FUNCTION_BLOCK "FB_ZonePID"
TITLE = Split-range heat/cool PID for one TCU zone
{ S7_Optimized_Access := 'TRUE' }
AUTHOR : chad416
VERSION : 0.2
//  Call every CycleTime seconds from a cyclic interrupt OB (e.g. OB30, 100 ms).
//  Output is in heating-equivalent percent: Output > 0 heats, Output < 0 cools.
//  CoolGainRatio = Kcool / Kheat (process gains). The cooling output is divided
//  by it so the loop gain is the same in both ranges.
//  FeedForward (heating-equivalent %) is added to the PID sum, through a
//  first-order lag FfTime (s); e.g. -FfGain * measured process power.
//  The float32 reference model is src/tcutune/pid.py: keep both in step.
   VAR_INPUT
      Setpoint : Real;   // degC
      Input : Real;   // measured temperature, degC
      ManualEnable : Bool;   // TRUE: Output := ManualValue (bumpless back to auto)
      ManualValue : Real;   // %, heating-equivalent
      Reset : Bool;   // clears integral and derivative state, outputs 0
      Gain : Real := 5.0;   // %/K
      Ti : Real := 300.0;   // s, 0 = no integral action
      Td : Real := 0.0;   // s, 0 = no derivative action
      DerivFilterN : Real := 10.0;   // derivative filter time constant = Td / N
      SpWeight : Real := 1.0;   // setpoint weight of the P part (0..1)
      Tt : Real := 0.0;   // s, anti-windup tracking time, <= 0 uses Ti
      CoolGainRatio : Real := 1.0;   // Kcool / Kheat
      Deadband : Real := 0.0;   // %, |Output| below this switches both actuators off
      CycleTime : Real := 0.1;   // s, call interval of the OB
      FeedForward : Real;   // %, heating-equivalent, 0 = none
      FfTime : Real := 0.0;   // s, lag on FeedForward, 0 = none
      CoolSaturated : Bool;   // FB_CoolLinearise.Saturated (last cycle): stop integrating into cooling
   END_VAR

   VAR_OUTPUT
      OutHeat : Real;   // % heater
      OutCool : Real;   // % cooling valve
      Output : Real;   // %, heating-equivalent controller output
   END_VAR

   VAR
      sI : Real;   // integral part
      sD : Real;   // filtered derivative part
      sPvPrev : Real;
      sF : Real;   // lagged feedforward
      sInitialised : Bool;
   END_VAR

   VAR_TEMP
      tP : Real;
      tA : Real;
      tU0 : Real;
      tU : Real;
      tOutLo : Real;
      tRatio : Real;
      tTt : Real;
      tInc : Real;
   END_VAR


BEGIN
	REGION Reset
	    IF #Reset THEN
	        #sI := 0.0;
	        #sD := 0.0;
	        #sF := 0.0;
	        #sInitialised := FALSE;
	        #Output := 0.0;
	        #OutHeat := 0.0;
	        #OutCool := 0.0;
	        RETURN;
	    END_IF;
	    IF NOT #sInitialised THEN
	        #sPvPrev := #Input;
	        #sF := #FeedForward;
	        #sInitialised := TRUE;
	    END_IF;
	END_REGION

	REGION Parameters
	    #tRatio := #CoolGainRatio;
	    IF #tRatio < 0.01 THEN
	        #tRatio := 0.01;
	    END_IF;
	    #tOutLo := -100.0 * #tRatio;
	    #tTt := #Tt;
	    IF #tTt <= 0.0 THEN
	        #tTt := #Ti;
	    END_IF;
	END_REGION

	REGION PID
	    #tP := #Gain * (#SpWeight * #Setpoint - #Input);

	    // derivative on the measurement, first-order filter, backward Euler
	    IF #Td > 0.0 THEN
	        #tA := #Td / (#Td + #DerivFilterN * #CycleTime);
	        #sD := #tA * #sD - #Gain * #DerivFilterN * #tA * (#Input - #sPvPrev);
	    ELSE
	        #sD := 0.0;
	    END_IF;

	    IF #FfTime > 0.0 THEN
	        #sF := #sF + #CycleTime / (#FfTime + #CycleTime) * (#FeedForward - #sF);
	    ELSE
	        #sF := #FeedForward;
	    END_IF;

	    #tU0 := #tP + #sI + #sD + #sF;

	    IF #ManualEnable THEN
	        #tU := LIMIT(MN := #tOutLo, IN := #ManualValue, MX := 100.0);
	        #sI := #tU - #tP - #sD - #sF;   // integral tracks the manual value
	    ELSE
	        #tU := LIMIT(MN := #tOutLo, IN := #tU0, MX := 100.0);
	        IF #Ti > 0.0 THEN
	            // integration plus back-calculation anti-windup
	            #tInc := #Gain * #CycleTime / #Ti * (#Setpoint - #Input);
	            IF #CoolSaturated AND #tU < 0.0 AND #tInc < 0.0 THEN
	                #tInc := 0.0;   // conditional integration: valve already fully open
	            END_IF;
	            #sI := #sI + #tInc + #CycleTime / #tTt * (#tU - #tU0);
	        ELSE
	            #sI := 0.0;
	        END_IF;
	    END_IF;
	END_REGION

	REGION Split_range
	    IF #tU >= #Deadband THEN
	        #OutHeat := #tU;
	        #OutCool := 0.0;
	    ELSIF #tU <= -#Deadband THEN
	        #OutHeat := 0.0;
	        #OutCool := MIN(IN1 := -#tU / #tRatio, IN2 := 100.0);
	    ELSE
	        #OutHeat := 0.0;
	        #OutCool := 0.0;
	    END_IF;
	    #Output := #tU;
	    #sPvPrev := #Input;
	END_REGION

END_FUNCTION_BLOCK
